// TIA Portal V21 export
// export: Created 2026-11-09T18:40:55.7554086Z, ExportSetting WithDefaults, DisplayName Totally Integrated Automation Portal, DisplayVersion V21 Update 3, DisplayName STEP 7 Professional, DisplayVersion V21 Update 3, DisplayName STEP 7 Safety, DisplayVersion V21, DisplayName Tech WebApplication, DisplayVersion V21, DisplayName WinCC Basic/Comfort/Advanced, DisplayVersion V21 Update 3, DisplayName WinCC Unified, DisplayVersion V21 Update 3
FUNCTION_BLOCK "FB_Lad_ex134"   // FB1, LAD
{ S7_Optimized_Access := 'TRUE' }
VERSION : 0.1
// stored: AutoNumber true, IsIECCheckEnabled false, IsRetainMemResEnabled false, MemoryReserve 100, SetENOAutomatically false, UDAEnableTagReadback false
   VAR_INPUT
      v_pwm : HW_PWM;
      v_enable : Bool;
   END_VAR
   VAR_OUTPUT
      v_busy : Bool;
      v_status : Word;
   END_VAR
   VAR
      inst { S7_SetPoint := 'True'} : CTRL_PWM;
   END_VAR
BEGIN

REGION Network 1: CTRL_PWM - Pulse-width modulation
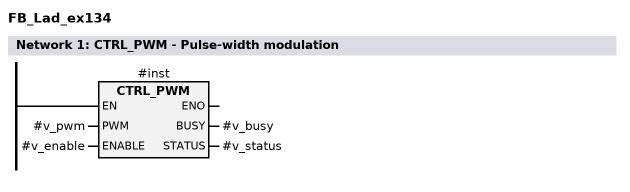
   RUNG wire#powerrail
      #inst.CTRL_PWM(PWM := #v_pwm, ENABLE := #v_enable, BUSY => #v_busy, STATUS => #v_status)
   END_RUNG
   // the same network as SCL:
   #inst(PWM := #v_pwm, ENABLE := #v_enable, BUSY => #v_busy, STATUS => #v_status);   // CTRL_PWM
END_REGION
END_FUNCTION_BLOCK
